Yaskawa INFORM job: HAND_OPEN.JBI

/JOB
//NAME HAND_OPEN
//POS
///NPOS 0,0,0,0,0,0
//INST
///DATE 2026/10/09 19:37
///COMM GRIPPER OPEN
///ATTR SC,RW
NOP
DOUT OT#(1) OFF
DOUT OT#(2) ON
WAIT IN#(2)=ON T=3.00
TIMER T=0.20
DOUT OT#(2) OFF
END
